PROGRAM main
  VAR
    B1 AT %IX0.0  : BOOL; (* sensor de piezas *)
    S1 AT %IX0.1  : BOOL; (* RESET *)
    KM1 AT %QX0.0 : BOOL; (* motor de la cinta *)
    H1 AT %QX0.1  : BOOL; (* aviso *)
    PIEZAS        : CTU;
    CUENTA        : INT; (* piezas en la caja *)
  END_VAR
  VAR  (* added by the conversion: wires and edge detectors of the diagram *)
    _LT6_OUT : BOOL;
    _GE10_OUT : BOOL;
  END_VAR

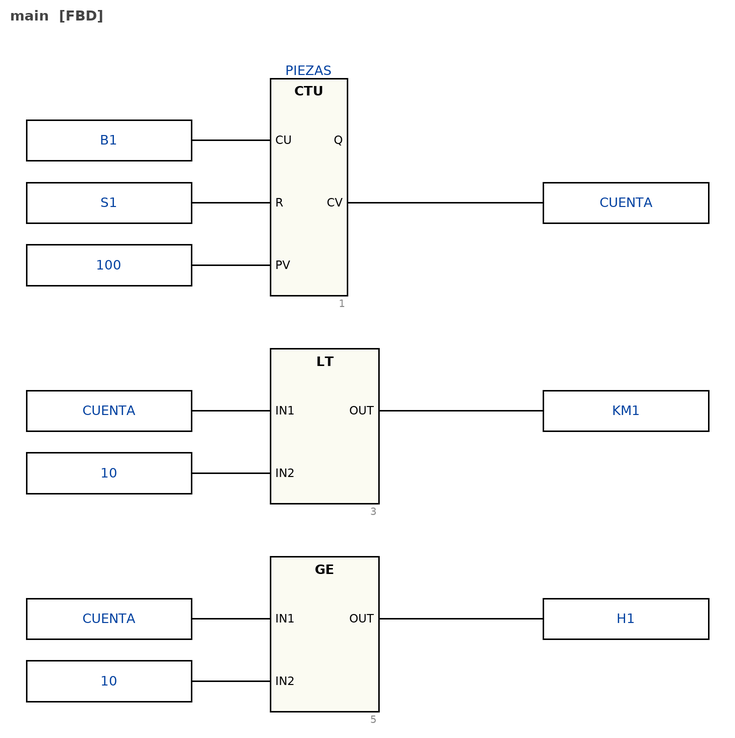
(* FBD diagram, written out as Structured Text *)
PIEZAS(CU := B1, R := S1, PV := 100);
CUENTA := PIEZAS.CV;
_LT6_OUT := CUENTA < 10;
KM1 := _LT6_OUT;
_GE10_OUT := CUENTA >= 10;
H1 := _GE10_OUT;
END_PROGRAM
